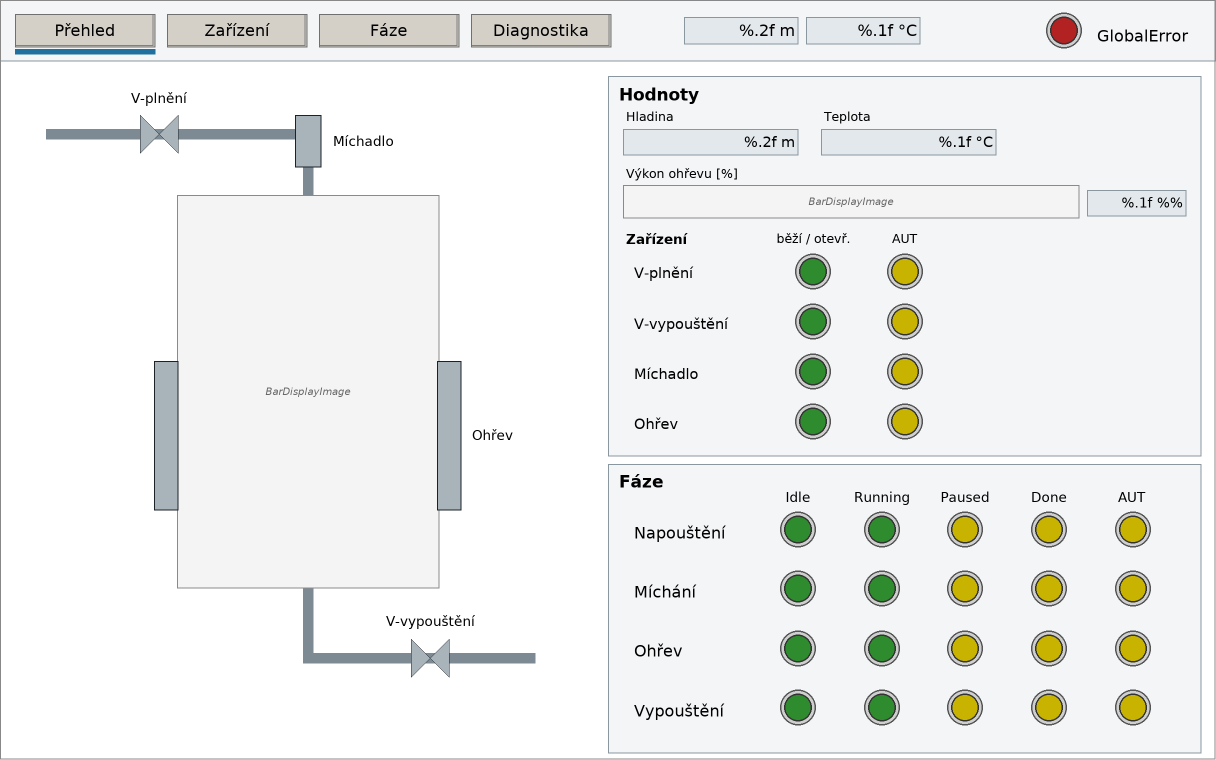
VISUALIZATION Prehled  // 1216x760
    Rectangle (0,0 1216x61)
    Button (15,14 140x33), "Přehled"
        OnMouseClick: change screen: Prehled
    Rectangle (15,49 140x5)
    Button (167,14 140x33), "Zařízení"
        OnMouseClick: change screen: Zarizeni
    Button (319,14 140x33), "Fáze"
        OnMouseClick: change screen: Faze
    Button (471,14 140x33), "Diagnostika"
        OnMouseClick: change screen: Diagnostika
    Rectangle (684,17 114x27), "%.2f m", text variable: Global.Tank1.Filling.WaterLevel
    Rectangle (806,17 114x27), "%.1f °C", text variable: Global.Tank1.Heating.WaterTemp
    Lamp1 (1041,10 46x41), variable: Global.Tank1.GlobalError, style: Lamp-Lamp1-Red
    Label (1094,23 126x26), "GlobalError"
    Rectangle (46,129 267x10)
    Rectangle (303,129 10x68)
    Rectangle (303,586 10x77)
    Rectangle (303,653 232x10)
    BarDisplayImage (177,195 262x393), value: Global.Tank1.Filling.WaterLevel, style: BarDisplayImage-Gray, scale format: %.1f, scale 0..2
    Polygon (140,115) (178,153) (178,115) (140,153) (140,153), colour toggle: Global.Tank1.ValveFilling.State.Open
    Label (121,87 76x23), "V-plnění"
    Polygon (411,639) (449,677) (449,639) (411,677) (411,677), colour toggle: Global.Tank1.ValveDraining.State.Open
    Label (385,610 91x23), "V-vypouštění"
    Rectangle (295,115 26x52), colour toggle: Global.Tank1.Mixer.State.Run
    Label (330,130 80x23), "Míchadlo"
    Rectangle (154,361 24x149), colour toggle: Global.Tank1.Heater.State.EnableOut
    Rectangle (437,361 24x149), colour toggle: Global.Tank1.Heater.State.EnableOut
    Label (469,424 52x23), "Ohřev"
    Rectangle (608,76 593x380)
    Label (616,81 87x27), "Hodnoty"
    Label (623,106 66x21), "Hladina"
    Rectangle (623,129 175x26), "%.2f m", text variable: Global.Tank1.Filling.WaterLevel
    Label (821,106 66x21), "Teplota"
    Rectangle (821,129 175x26), "%.1f °C", text variable: Global.Tank1.Heating.WaterTemp
    Label (623,163 142x21), "Výkon ohřevu [%]"
    BarDisplayImage (623,185 456x33), value: Global.Tank1.Heater.State.HeatingOut, style: BarDisplayImage-Gray, scale format: %.1f, scale 0..100
    Rectangle (1087,190 99x26), "%.1f %%", text variable: Global.Tank1.Heater.State.HeatingOut
    Label (623,228 80x23), "Zařízení"
    Label (768,228 91x21), "běží / otevř."
    Label (859,228 91x21), "AUT"
    Label (631,261 84x24), "V-plnění"
    Lamp1 (790,251 46x41), variable: Global.Tank1.ValveFilling.State.Open, style: Lamp-Lamp1-Green
    Lamp1 (882,251 46x41), variable: Global.Tank1.ValveFilling.State.AutCtrl, style: Lamp-Lamp1-Yellow
    Label (631,312 123x24), "V-vypouštění"
    Lamp1 (790,301 46x41), variable: Global.Tank1.ValveDraining.State.Open, style: Lamp-Lamp1-Green
    Lamp1 (882,301 46x41), variable: Global.Tank1.ValveDraining.State.AutCtrl, style: Lamp-Lamp1-Yellow
    Label (631,362 84x24), "Míchadlo"
    Lamp1 (790,351 46x41), variable: Global.Tank1.Mixer.State.Run, style: Lamp-Lamp1-Green
    Lamp1 (882,351 46x41), variable: Global.Tank1.Mixer.State.AutCtrl, style: Lamp-Lamp1-Yellow
    Label (631,412 55x24), "Ohřev"
    Lamp1 (790,401 46x41), variable: Global.Tank1.Heater.State.EnableOut, style: Lamp-Lamp1-Green
    Lamp1 (882,401 46x41), variable: Global.Tank1.Heater.State.AutCtrl, style: Lamp-Lamp1-Yellow
    Rectangle (608,464 593x289)
    Label (616,468 53x27), "Fáze"
    Label (760,486 76x23), "Idle"
    Label (844,486 76x23), "Running"
    Label (927,486 76x23), "Paused"
    Label (1011,486 76x23), "Done"
    Label (1094,486 76x23), "AUT"
    Label (631,520 116x26), "Napouštění"
    Lamp1 (775,509 46x41), variable: Global.Tank1.Filling.State.Idle, style: Lamp-Lamp1-Green
    Lamp1 (859,509 46x41), variable: Global.Tank1.Filling.State.Running, style: Lamp-Lamp1-Green
    Lamp1 (942,509 46x41), variable: Global.Tank1.Filling.State.Paused, style: Lamp-Lamp1-Yellow
    Lamp1 (1026,509 46x41), variable: Global.Tank1.Filling.State.Done, style: Lamp-Lamp1-Yellow
    Lamp1 (1110,509 46x41), variable: Global.Tank1.Filling.State.AutCtrl, style: Lamp-Lamp1-Yellow
    Label (631,579 83x26), "Míchání"
    Lamp1 (775,568 46x41), variable: Global.Tank1.Mixing.State.Idle, style: Lamp-Lamp1-Green
    Lamp1 (859,568 46x41), variable: Global.Tank1.Mixing.State.Running, style: Lamp-Lamp1-Green
    Lamp1 (942,568 46x41), variable: Global.Tank1.Mixing.State.Paused, style: Lamp-Lamp1-Yellow
    Lamp1 (1026,568 46x41), variable: Global.Tank1.Mixing.State.Done, style: Lamp-Lamp1-Yellow
    Lamp1 (1110,568 46x41), variable: Global.Tank1.Mixing.State.AutCtrl, style: Lamp-Lamp1-Yellow
    Label (631,638 62x26), "Ohřev"
    Lamp1 (775,628 46x41), variable: Global.Tank1.Heating.State.Idle, style: Lamp-Lamp1-Green
    Lamp1 (859,628 46x41), variable: Global.Tank1.Heating.State.Running, style: Lamp-Lamp1-Green
    Lamp1 (942,628 46x41), variable: Global.Tank1.Heating.State.Paused, style: Lamp-Lamp1-Yellow
    Lamp1 (1026,628 46x41), variable: Global.Tank1.Heating.State.Done, style: Lamp-Lamp1-Yellow
    Lamp1 (1110,628 46x41), variable: Global.Tank1.Heating.State.AutCtrl, style: Lamp-Lamp1-Yellow
    Label (631,698 116x26), "Vypouštění"
    Lamp1 (775,687 46x41), variable: Global.Tank1.Draining.State.Idle, style: Lamp-Lamp1-Green
    Lamp1 (859,687 46x41), variable: Global.Tank1.Draining.State.Running, style: Lamp-Lamp1-Green
    Lamp1 (942,687 46x41), variable: Global.Tank1.Draining.State.Paused, style: Lamp-Lamp1-Yellow
    Lamp1 (1026,687 46x41), variable: Global.Tank1.Draining.State.Done, style: Lamp-Lamp1-Yellow
    Lamp1 (1110,687 46x41), variable: Global.Tank1.Draining.State.AutCtrl, style: Lamp-Lamp1-Yellow
END_VISUALIZATION

(* stored: Version 1.1.0.1, ProductVersion 3.1.4024.16
   Visu Prehled: Id {d71dcd47-18b0-43a6-a3d5-60ed4d052581} *)
